// TIA Portal project "LAB03" (V16)

(* hardware
DEVICE "S7300/ET200M station_1"  S7-300 station
   slot 0: "Rail_0"  Rail  6ES7 390-1***0-0AA0
   slot 1: "PS 307 2A_1"  PS 307 2A  6ES7 307-1BA00-0AA0
   slot 2: "PLC_1"  CPU 313C-2 DP  6ES7 313-6CF03-0AB0  V2.6
      slot 0: "MPI interface_1"  X1
      slot 1: "DP interface_1"  X2
      slot 2: "DI 16/DO 16_1"  DI16/DO16
      slot 4: "Count_1"  Counter
*)

// ===== PLC "PLC_1"  CPU 313C-2 DP =====

VAR_GLOBAL   // PLC tag table "Default tag table"
   "Tag_1" AT %Z5 : Counter;
   "Tag_2" AT %MW10 : Word;
END_VAR

DATA_BLOCK "DB10"   // DB10
{ S7_Optimized_Access := 'FALSE' }
VERSION : 0.1
   VAR
      Static_1 : DInt;
      Static_2 : DInt;
      Static_3 : DInt;
      Static_4 : DInt;
      Static_5 : DInt;
      Static_6 : DInt;
      Static_7 : DInt;
      Static_8 : DInt;
      Static_9 : DInt;
      Static_10 : DInt;
      Static_11 : DInt;
      Static_12 : DInt;
      Static_13 : DInt;
      Static_14 : DInt;
      Static_15 : DInt;
      Static_16 : DInt;
   END_VAR
BEGIN
END_DATA_BLOCK

FUNCTION "FC5" : Void   // FC5, STL
{ S7_Optimized_Access := 'FALSE' }
VERSION : 0.1
BEGIN

REGION Network 1
         A     %DB10.DBX1.0;  // if acquisition error
         =     %DB10.DBX8.0;  // copy on error bit, write FFFF on DBW6 and return
         JC    FAUL;
         L     %DB10.DBW0;  // load the acquired bit pattern
         SLW   3;  // shift left 3 bits
         SRW   4;  // shift right 4 bits
         T     "Tag_2";  // save in MW10
         L     %DB10.DBW2;  // load high threshold
         >I;  // check if value greater than threshold
         =     %DB10.DBX8.1;  // copy result of comparison on bit 8.1
         L     %DB10.DBW4;  // load low threshold
         L     "Tag_2";  // load value
         >I;  // check if value less than threshold
         =     %DB10.DBX8.2;  // copy result of comparison on bit 8.2
         O     %DB10.DBX8.1;  // if a threshold has been overcome
         O     %DB10.DBX8.2;
         JC    FAUL;  // write FFFF on DBW6 and return
         L     "Tag_2";  // else copy value on DB
         T     %DB10.DBW6;
         BEU;
   FAUL: L     w#16#ffff;  // error section: write ffff on DBW6
         T     %DB10.DBW6;
END_REGION
END_FUNCTION

FUNCTION "FC51" : Void   // FC51, STL
{ S7_Optimized_Access := 'FALSE' }
VERSION : 0.1
BEGIN

REGION Network 1
         A     %DB10.DBX1.0;  // if acquisition error
         =     %DB10.DBX8.0;  // copy on error bit, write FFFF on DBW6 and return
         JC    FAUL;
         L     %DB10.DBW0;  // load the acquired bit pattern
         SLW   3;  // shift left 3 bits
         SRW   4;  // shift right 4 bits
         T     "Tag_2";  // save in MW10
         L     %DB10.DBW2;  // load high threshold
         >I;  // check if value greater than threshold
         =     %DB10.DBX8.1;  // copy result of comparison on bit 8.1
         L     %DB10.DBW4;  // load low threshold
         L     "Tag_2";  // load value
         >I;  // check if value less than threshold
         =     %DB10.DBX8.2;  // copy result of comparison on bit 8.2
         L     "Tag_2";  // save value of
         L     %DB10.DBW12;  // load HIGH Warning
         >I;  //
         =     %DB10.DBX8.3;
         L     %DB10.DBW14;
         L     "Tag_2";  // save value of
         >I;
         =     %DB10.DBX8.4;
         O     %DB10.DBX8.1;  // if a threshold has been overcome
         O     %DB10.DBX8.2;
         O     %DB10.DBX8.3;  // if a threshold has been overcome
         O     %DB10.DBX8.4;
         =     %DB10.DBX8.7;
         O     %DB10.DBX8.1;  // if a threshold has been overcome
         O     %DB10.DBX8.2;
         JC    FAUL;  // write FFFF on DBW6 and return
         L     "Tag_2";  // else copy value on DB
         T     %DB10.DBW6;
         BEU;
   FAUL: L     w#16#ffff;  // error section: write ffff on DBW6
         T     %DB10.DBW6;
END_REGION
END_FUNCTION

ORGANIZATION_BLOCK "Main"   // OB1, STL
TITLE = "Main Program Sweep (Cycle)"
{ S7_Optimized_Access := 'FALSE' }
VERSION : 0.1
   VAR_TEMP
      OB1_EV_CLASS : Byte;   // Bits 0-3 = 1 (Coming event), Bits 4-7 = 1 (Event class 1)
      OB1_SCAN_1 : Byte;   // 1 (Cold restart scan 1 of OB 1), 3 (Scan 2-n of OB 1)
      OB1_PRIORITY : Byte;   // Priority of OB Execution
      OB1_OB_NUMBR : Byte;   // 1 (Organization block 1, OB1)
      OB1_RESERVED_1 : Byte;   // Reserved for system
      OB1_RESERVED_2 : Byte;   // Reserved for system
      OB1_PREV_CYCLE : Int;   // Cycle time of previous OB1 scan (milliseconds)
      OB1_MIN_CYCLE : Int;   // Minimum cycle time of OB1 (milliseconds)
      OB1_MAX_CYCLE : Int;   // Maximum cycle time of OB1 (milliseconds)
      OB1_DATE_TIME : Date_And_Time;   // Date and time OB1 started
   END_VAR
BEGIN

REGION Network 1
         CALL  "FC5";
END_REGION
END_ORGANIZATION_BLOCK